(* PLC project zarechnaya.project, CODESYS CODESYS V3.5 SP17 Patch 3 *)
(* stored: creationDateTime 2026-10-20T05:42:22.2197262, modificationDateTime 1601-01-01T03:00:00 *)

(* PRG_Permissives — разрешения пуска насоса промывки (LD, PROGRAM: P/N, S/R). Поведение (модель scenarios/reference/model_PRG_Permissives.py): 1. фронт xStartBtn И xPermit → xRun := TRUE (S); 2. спад xStopBtn ИЛИ NOT xPermit → xRun := FALSE (R) — сеть 2 после сети 1, сброс побеждает в одном цикле; 3. xMotor := xRun AND NOT xFault; 4. xIdle := NOT xRun (инверсная катушка). Фронты — R_TRIG/F_TRIG CODESYS по переменной; первый вызов: память фронта FALSE. *)
PROGRAM PRG_Permissives
  VAR_INPUT
    xStartBtn : BOOL;
    xStopBtn : BOOL;
    xPermit : BOOL;
    xFault : BOOL;
  END_VAR
  VAR_OUTPUT
    xRun : BOOL;
    xMotor : BOOL;
    xIdle : BOOL;
  END_VAR
  VAR  (* added by the conversion: wires and edge detectors of the diagram *)
    R_TRIG1 : R_TRIG;
    F_TRIG2 : F_TRIG;
  END_VAR

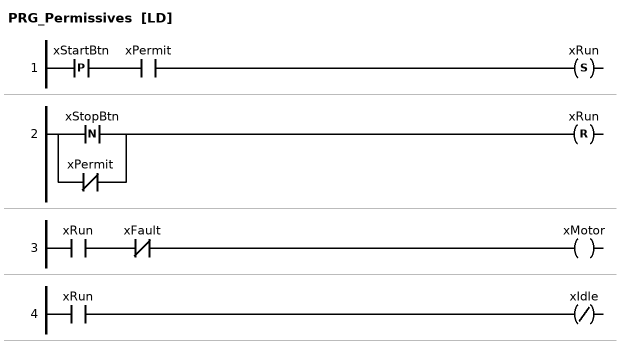
(* LD diagram, written out as Structured Text *)
(* --- network: Пуск по фронту --- *)
R_TRIG1(CLK := xStartBtn);
IF R_TRIG1.Q AND xPermit THEN xRun := TRUE; END_IF;
(* --- network: Стоп по спаду или без разрешения --- *)
F_TRIG2(CLK := xStopBtn);
IF F_TRIG2.Q OR NOT xPermit THEN xRun := FALSE; END_IF;
(* --- network: Двигатель --- *)
xMotor := xRun AND NOT xFault;
(* --- network: Простой --- *)
xIdle := NOT xRun;
END_PROGRAM
